{attribute 'no_assign'}
FUNCTION_BLOCK FB_LN_WTURBINE_LD0_WYAW1 EXTENDS FB_AcsiCommonLogicalNodeClass
VAR_INPUT
	Beh: FB_DO_WTURBINE_LD0_WYAW1_Beh := (sClass:='ENS', bLinkResult:=THIS^.AddDataToContainer(ipData:=Beh));
	YwAng: FB_DO_WTURBINE_LD0_WYAW1_YwAng := (sClass:='MV', bLinkResult:=THIS^.AddDataToContainer(ipData:=YwAng));
	CabWup: FB_DO_WTURBINE_LD0_WYAW1_CabWup := (sClass:='MV', bLinkResult:=THIS^.AddDataToContainer(ipData:=CabWup));
	YwAngSpt: FB_DO_WTURBINE_LD0_WYAW1_YwAngSpt := (sClass:='SPV', bLinkResult:=THIS^.AddDataToContainer(ipData:=YwAngSpt));
END_VAR
VAR
END_VAR

END_FUNCTION_BLOCK

(* stored: Version 1.1.0.1
   POU FB_LN_WTURBINE_LD0_WYAW1: Id {4ea6dc1f-8b13-49c3-9d45-dc4cc3d5423a}, SpecialFunc None *)
